Fanuc KAREL source: ka00065.KL

-- PROVISIONAL review KL for V1013-1; original PC SHA256 d771a3a55cd5bc89ba9394f2bf305502fcb304811c115681bfc4cf9b8ecf81bc
-- Incomplete behavior may be omitted. Consult companion uncertainty JSON. Do not deploy.
PROGRAM KA00065
%NOLOCKGROUP
-- UNRESOLVED_DECL SRC type=000102
-- UNRESOLVED_DECL DST type=000101
BEGIN
  -- UNRESOLVED_PC offsets 5-20; opcodes 2E,22,32,35
  -- UNRESOLVED_PC offsets 25-45; opcodes 49,7E,4A
  -- UNRESOLVED_PC offsets 50-54; opcodes 7F
END KA00065
